// TIA Portal V19 export
// export: Created 2026-10-15T10:10:36.8885543Z, ExportSetting WithDefaults, DisplayName Totally Integrated Automation Portal, DisplayVersion V19, DisplayName TIA Portal Openness, DisplayVersion V19, DisplayName TIA Portal Version Control Interface, DisplayVersion V19, DisplayName STEP 7 Professional, DisplayVersion V19, DisplayName STEP 7 Safety, DisplayVersion V19, DisplayName WinCC Basic/Comfort/Advanced, DisplayVersion V19, DisplayName WinCC Unified, DisplayVersion V19
FUNCTION "ROLL_PB24" : Void   // FC31, SCL
{ S7_Optimized_Access := 'TRUE' }
VERSION : 0.1
// stored: AutoNumber true, IsIECCheckEnabled false, SetENOAutomatically false, UDAEnableTagReadback false
   VAR_TEMP
      r : Bool;
      a1 : Word;
      a2 : Word;
      activeDataBlock : Int;
      comparisonResults : Array[0..0] of Bool;
   END_VAR
BEGIN

   #r := FALSE;
   #a1 := W#16#0000;
   #a2 := W#16#0000;
   #activeDataBlock := 0;
   // PB24, STEP 5 network 1
   #activeDataBlock := 15;
   // PB24, STEP 5 network 2
   #r := ("ROLL_IO".Input[5, 0] AND "ROLL_State".M[13, 3] AND "ROLL_State".S5Timers[59].Q);
   "ROLL_State".M[240, 0] := #r;
   // PB24, STEP 5 network 3
   #a2 := #a1;
   #a1 := "ROLL_GetDW"(DbNumber := #activeDataBlock, Index := 54);
   #r := (NOT "ROLL_State".S5Timers[53].Q);
   "ROLL_TimerOp"(Number := 54,
                  Operation := 0,
                  Signal := #r,
                  Preset := #a1);
   #a2 := #a1;
   #a1 := "ROLL_GetDW"(DbNumber := #activeDataBlock, Index := 53);
   #r := "ROLL_State".S5Timers[54].Q;
   "ROLL_TimerOp"(Number := 53,
                  Operation := 1,
                  Signal := #r,
                  Preset := #a1);
   #r := "ROLL_State".M[240, 0];
   "ROLL_TimerOp"(Number := 53,
                  Operation := 2,
                  Signal := #r,
                  Preset := #a1);
   #r := ((NOT "ROLL_State".M[40, 5]) AND "ROLL_State".S5Timers[53].Q);
   "ROLL_IO".Output[19, 4] := #r;
   // PB24, STEP 5 network 4
   RETURN;
END_FUNCTION
